PROGRAM Gr01MachineMode
VAR_INPUT
	(* Input variables / Eingang Variablen *)
	bEnable					:BOOL;						(* Enable Gr01MachineMode *)
END_VAR
VAR
	(* Enummerations *)

	(* Variables *)

	(* References *)

	(* Interfaces *)

	(* Instances *)

END_VAR

IF NOT bEnable
THEN
	RETURN;
END_IF;

Gr01Auto(bEnable := TRUE);			(* Call Program *)
Gr01Home(bEnable := TRUE);			(* Call Program *)
Gr01Manual(bEnable := TRUE);			(* Call Program *)

END_PROGRAM

(* stored: Version 1.1.0.1, ProductVersion 3.1.4024.15
   POU Gr01MachineMode: Id {ac484db5-f68a-43dc-91fe-db60cf5f173f}, SpecialFunc None *)
